Staubli VAL3: bind.pgx

program bind()
  local num l_i
  local string l_sbtn
begin
  //lbllib
  userPageBind("traj","lbllib","innerHTML",sUsingLib,1,"r")
  //lst
  //  if size(sList)<50
  //    userPageBind("traj","lst1","options",sList,size(sList),"r")
  //    else
  //      popUpMsg("traj数量过大")
  //    endIf
  userPageBind("traj","lst1","value",sSelTraj,1,"rw")
  //button
  userPageBindClick("traj","btnback",bBack,true)
  for l_i = 0 to 11
    l_sbtn="btn"+toString("",l_i)
    userPageBindClick("traj",l_sbtn,bBool[l_i],true)
  endFor

  //page
  userPageBind("traj","lblpageindex","innerHTML",sPageIndex,1,"r")

  userPageBind("traj","lblpagenum","innerHTML",sPageNum,1,"r")


end
